// LS Electric XG5000 project: error-reset
// PLC LSPLC

PROGRAM error-reset (task: 스캔 프로그램)

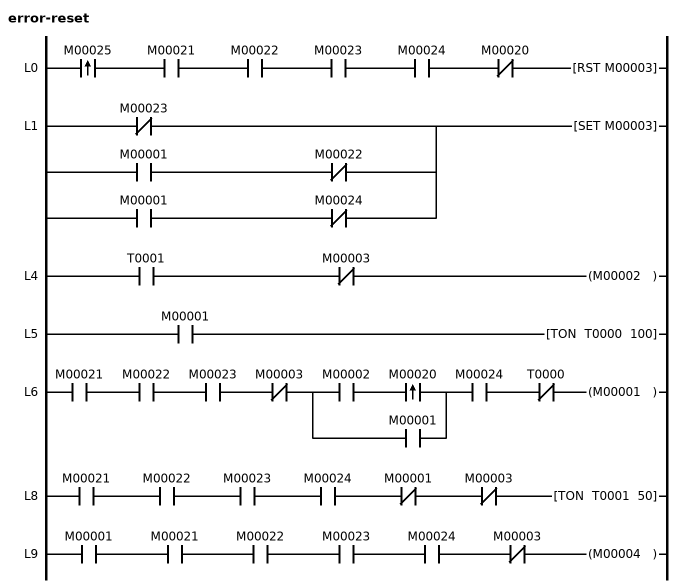
; L0
LOADP     M00025
AND       M00021
AND       M00022
AND       M00023
AND       M00024
AND NOT   M00020
RST       M00003
; L1
LOAD NOT  M00023
LOAD      M00001
AND NOT   M00022
OR LOAD
LOAD      M00001
AND NOT   M00024
OR LOAD
SET       M00003
; L4
LOAD      T0001
AND NOT   M00003
OUT       M00002
; L5
LOAD      M00001
TON       T0000 100
; L6
LOAD      M00021
AND       M00022
AND       M00023
AND NOT   M00003
LOAD      M00002
ANDP      M00020
OR        M00001
AND LOAD
AND       M00024
AND NOT   T0000
OUT       M00001
; L8
LOAD      M00021
AND       M00022
AND       M00023
AND       M00024
AND NOT   M00001
AND NOT   M00003
TON       T0001 50
; L9
LOAD      M00001
AND       M00021
AND       M00022
AND       M00023
AND       M00024
AND NOT   M00003
OUT       M00004